Fanuc KAREL source: kt00409.KL

PROGRAM KT00409
%NOLOCKGROUP
VAR
B1:BOOLEAN;B2:BOOLEAN;OUT:BOOLEAN
BEGIN
--
--
B1=TRUE
B2=FALSE
B1=TRUE
B2=FALSE
OUT=(B1>B2)
END KT00409
